// TIA Portal V21 export
// export: Created 2026-08-21T20:18:52.0347368Z, ExportSetting None, DisplayName Totally Integrated Automation Portal, DisplayVersion V21, DisplayName STEP 7 Professional, DisplayVersion V21, DisplayName STEP 7 Safety, DisplayVersion V21, DisplayName Tech WebApplication, DisplayVersion V21, DisplayName WinCC Basic/Comfort/Advanced, DisplayVersion V21, DisplayName WinCC Professional, DisplayVersion V21, DisplayName WinCC Unified, DisplayVersion V21
DATA_BLOCK "CMInterface_DB"   // DB27
// stored: InstanceOfName CM_Interface, InstanceOfType FB
"CM_Interface"
   // VAR_INPUT
   //    CmCommand { ExternalAccessible := 'False'; ExternalVisible := 'False'; ExternalWritable := 'False'} : Array[0..29] of Bool;
   //    Procedure_Param { ExternalAccessible := 'False'; ExternalVisible := 'False'; ExternalWritable := 'False'} : Array[0..31] of Real;
   //    Config_Param : Array[0..31] of Bool;
   //    ProcessValueIn_Bool : Array[0..31] of Bool;
   //    ProcessValueIn_Real : Array[0..31] of Real;
   //    CmFbOnOff { ExternalAccessible := 'False'; ExternalVisible := 'False'; ExternalWritable := 'False'} : Array[0..29] of Bool;
   //    DosingSpeed : Real;
   //    Auto_Man : Bool;
   //    Oos : Bool;
   // END_VAR
   // VAR_OUTPUT
   //    CM_P100 { ExternalAccessible := 'False'; ExternalVisible := 'False'; ExternalWritable := 'False'} : "DigVal";
   //    CM_P101 { ExternalAccessible := 'False'; ExternalVisible := 'False'; ExternalWritable := 'False'} : "DigVal";
   //    CM_FIC100 { ExternalAccessible := 'False'; ExternalVisible := 'False'; ExternalWritable := 'False'} : "DigVal";
   //    CM_V100 { ExternalAccessible := 'False'; ExternalVisible := 'False'; ExternalWritable := 'False'} : "DigVal";
   //    FlowRate { ExternalAccessible := 'False'; ExternalVisible := 'False'; ExternalWritable := 'False'} : "AnaVal";
   //    Liter { ExternalAccessible := 'False'; ExternalVisible := 'False'; ExternalWritable := 'False'} : "AnaVal";
   //    ExternalLevel : "AnaVal";
   //    PEA_inlet_Vlv_opened : "DigVal";
   //    PVConnected : "DigVal";
   // END_VAR
   // VAR
   //    Pos_edge : Bool;
   //    Neg_edge : Bool;
   // END_VAR
BEGIN
END_DATA_BLOCK
